FUNCTION_BLOCK F (* Negative C3: a copy of a copy of the position, read by guards *)
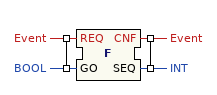
  EVENT_INPUT
    REQ WITH GO;
  END_EVENT
  EVENT_OUTPUT
    CNF WITH SEQ;
  END_EVENT
  VAR_INPUT
    GO : BOOL;
  END_VAR
  VAR_OUTPUT
    SEQ : INT;
  END_VAR
  VAR
    K : INT;
    L : INT;
  END_VAR
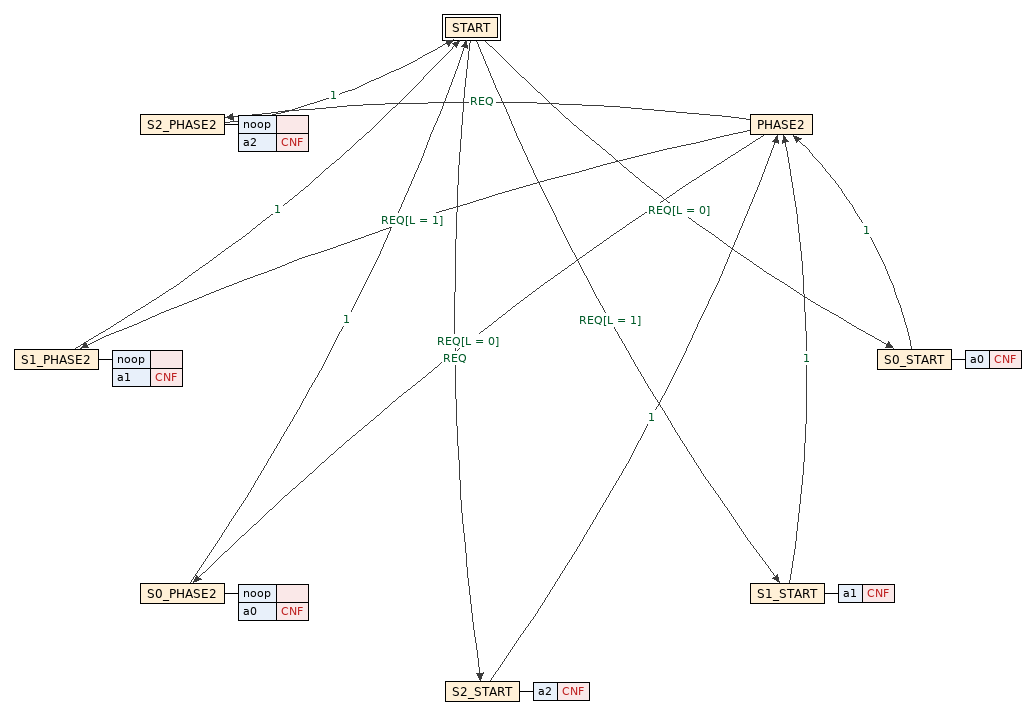
  EC_STATES
    START;
    PHASE2;
    S0_START : a0 -> CNF;
    S1_START : a1 -> CNF;
    S2_START : a2 -> CNF;
    S0_PHASE2 : noop, a0 -> CNF;
    S1_PHASE2 : noop, a1 -> CNF;
    S2_PHASE2 : noop, a2 -> CNF;
  END_STATES
  EC_TRANSITIONS
    START TO S0_START := REQ[L = 0];
    START TO S1_START := REQ[L = 1];
    START TO S2_START := REQ;
    PHASE2 TO S0_PHASE2 := REQ[L = 0];
    PHASE2 TO S1_PHASE2 := REQ[L = 1];
    PHASE2 TO S2_PHASE2 := REQ;
    S0_START TO PHASE2 := 1;
    S1_START TO PHASE2 := 1;
    S2_START TO PHASE2 := 1;
    S0_PHASE2 TO START := 1;
    S1_PHASE2 TO START := 1;
    S2_PHASE2 TO START := 1;
  END_TRANSITIONS
  ALGORITHM a0 IN ST:
IF GO THEN
  SEQ := 1;
END_IF;
K := SEQ;
L := K;
  END_ALGORITHM
  ALGORITHM a1 IN ST:
SEQ := 2;
K := SEQ;
L := K;
  END_ALGORITHM
  ALGORITHM a2 IN ST:
SEQ := 0;
K := SEQ;
L := K;
  END_ALGORITHM
  ALGORITHM noop IN ST:
K := K;
  END_ALGORITHM
END_FUNCTION_BLOCK
